(* IEC 61131-3 sources: ControlsBenchMUSE/codesys/library/source, 19 files *)

(* ---- ST_CB_Config.st ---- *)
TYPE ST_CB_Config :
STRUCT
    DomainId : UDINT; // nonzero; unique per authority domain in the application
    SchemaId : UDINT; // nonzero machine-map fingerprint of the raw channel layout
    TimeoutUs : ULINT := 500000; // heartbeat staleness as elapsed microseconds
    DigitalCount : UINT; // configured channels occupy indices 0..Count-1 of each bank
    SignedCount : UINT;
    UnsignedCount : UINT;
    RealCount : UINT;
    SignedBits : ARRAY[0..31] OF USINT; // native width of each configured channel: 8, 16 or 32
    UnsignedBits : ARRAY[0..31] OF USINT; // native width of each configured channel: 1 to 32
    RealNonFiniteAllowed : ARRAY[0..15] OF BOOL; // TRUE only where the device can report NaN or infinity
END_STRUCT
END_TYPE

(* ---- ST_CB_Image.st ---- *)
TYPE ST_CB_Image :
STRUCT
    Digital : ARRAY[0..63] OF BOOL;
    Numeric : ST_CB_Numeric;
END_STRUCT
END_TYPE

(* ---- ST_CB_ImageMask.st ---- *)
TYPE ST_CB_ImageMask :
STRUCT
    Digital : ARRAY[0..63] OF BOOL;
    Numeric : ST_CB_NumericMask;
END_STRUCT
END_TYPE

(* ---- ST_CB_Numeric.st ---- *)
TYPE ST_CB_Numeric :
STRUCT
    Signed : ARRAY[0..31] OF DINT;
    Unsigned : ARRAY[0..31] OF UDINT;
    RealValue : ARRAY[0..15] OF REAL;
END_STRUCT
END_TYPE

(* ---- ST_CB_NumericMask.st ---- *)
TYPE ST_CB_NumericMask :
STRUCT
    Signed : ARRAY[0..31] OF BOOL;
    Unsigned : ARRAY[0..31] OF BOOL;
    RealValue : ARRAY[0..15] OF BOOL;
END_STRUCT
END_TYPE

(* ---- ST_CB_ObservationFrame.st ---- *)
TYPE ST_CB_ObservationFrame :
STRUCT
    FrameFormat : UDINT := 1; // GVL_CB.FRAME_FORMAT_VERSION
    FrameSequence : ULINT; // frames published by this block since initialization
    BootIdentity : ULINT;
    DomainId : UDINT;
    SchemaId : UDINT;
    TapSchemaId : UDINT; // fingerprint of the configured tap list; 0 when none is configured
    SourceCycle : ULINT; // session cycle whose inputs and outputs this frame holds
    SourceTimeUs : ULINT; // platform monotonic time at capture, not wall-clock time
    CapturePhase : USINT; // GVL_CB.PHASE_POST_OUTPUT
    MissedCycles : ULINT; // cumulative session cycles that published no frame
    RepeatedCycles : ULINT; // cumulative calls without a new session cycle (integration error)
    SimApplied : BOOL; // SelectedInputs came from the workstation, not hardware
    ConnectorStale : BOOL;
    ConfigValid : BOOL;
    ClockValid : BOOL;
    ReconfigureRequired : BOOL;
    AnySuppressed : BOOL;
    AppliedEpoch : ULINT;
    AppliedSequence : ULINT;
    RawInputs : ST_CB_Image; // hardware values presented to the session, in either mode
    SelectedInputs : ST_CB_Image; // image the application consumed
    Commands : ST_CB_Image; // authentic application commands before suppression
    Physical : ST_CB_Image; // physical sink values after suppression
    Suppressed : ST_CB_ImageMask; // channels whose physical sink was suppressed
    Taps : ST_CB_Image; // explicitly configured observation taps; never writable through this library
END_STRUCT
END_TYPE

(* ---- ST_CB_Request.st ---- *)
TYPE ST_CB_Request :
STRUCT
    SimRequest : BOOL;
    SimulationResetRequest : BOOL; // rising edge: zero image, remain simulated
    SessionResetRequest : BOOL;
    Heartbeat : ULINT;
    RequestedSlot : USINT := 255;
    RequestedEpoch : ULINT;
    RequestedSequence : ULINT; // write LAST after validity/payload/metadata
    Slots : ARRAY[0..1] OF ST_CB_Slot;
END_STRUCT
END_TYPE

(* ---- ST_CB_Slot.st ---- *)
TYPE ST_CB_Slot :
STRUCT
    Valid : BOOL;
    DomainId : UDINT;
    SchemaId : UDINT;
    Epoch : ULINT;
    Sequence : ULINT;
    Data : ST_CB_Image;
END_STRUCT
END_TYPE

(* ---- ST_CB_Status.st ---- *)
TYPE ST_CB_Status :
STRUCT
    ProtocolVersion : UDINT := 2; // GVL_CB.PROTOCOL_VERSION
    DomainId : UDINT; // pinned at initialization
    SchemaId : UDINT; // pinned at initialization
    ConfigValid : BOOL;
    ClockValid : BOOL; // this cycle's time was not earlier than the previous cycle's
    ReconfigureRequired : BOOL; // latched by config, boot or clock change; cleared only by Reinitialize
    SimApplied : BOOL; // TRUE: the application consumes the workstation image
    ConnectorStale : BOOL := TRUE;
    BootIdentity : ULINT;
    Cycle : ULINT; // calls of this domain session, not universal PLC scans
    TimeUs : ULINT;
    LastHeartbeat : ULINT;
    LastHeartbeatTimeUs : ULINT;
    ActiveSlot : USINT := 255;
    AppliedEpoch : ULINT;
    AppliedSequence : ULINT;
    AppliedCycle : ULINT;
    AppliedTimeUs : ULINT;
    // Acknowledgement of the last consumed request event, accepted or not.
    ConsumedEpoch : ULINT;
    ConsumedSequence : ULINT;
    ConsumedSlot : USINT := 255;
    ConsumedResult : UINT; // GVL_CB.RESULT_*
    ConsumedCycle : ULINT;
    ConsumedTimeUs : ULINT;
    RejectBank : USINT; // GVL_CB.BANK_* of the first channel failing representation checks
    RejectIndex : UINT;
    CommitCount : ULINT;
    DuplicateCount : ULINT;
    StaleCount : ULINT;
    SkippedCount : ULINT;
    InvalidSlotCount : ULINT;
    IncompleteSlotCount : ULINT;
    MetadataMismatchCount : ULINT;
    RepresentationRejectedCount : ULINT;
    EpochRejectedCount : ULINT;
    NotSimulatedCount : ULINT;
    BlockedRequestCount : ULINT;
    IdleClearCount : ULINT;
    SessionResetCount : ULINT;
    SimulationResetCount : ULINT;
    SimulationEntryCount : ULINT;
    ReinitializeCount : ULINT;
END_STRUCT
END_TYPE

(* ---- U_CB_Real32.st ---- *)
TYPE U_CB_Real32 :
UNION
    AsReal : REAL; // IEEE 754 binary32 value
    AsBits : DWORD; // the same 32 bits, for encoding checks without numeric conversion
END_UNION
END_TYPE

(* ---- GVL_CB.st ---- *)
{attribute 'qualified_only'}
VAR_GLOBAL CONSTANT
    // Interface versions. The package version is the library project version (VERSIONING.md).
    API_VERSION_MAJOR : UINT := 0;
    API_VERSION_MINOR : UINT := 2;
    PROTOCOL_VERSION : UDINT := 2; // request, slot and status semantics of this raw-bank profile
    FRAME_FORMAT_VERSION : UDINT := 1; // ST_CB_ObservationFrame layout and meaning
    // Fixed capacities of ST_CB_Image. Configured channels occupy indices 0..Count-1.
    DIGITAL_CAPACITY : UINT := 64;
    SIGNED_CAPACITY : UINT := 32;
    UNSIGNED_CAPACITY : UINT := 32;
    REAL_CAPACITY : UINT := 16;
    NO_SLOT : USINT := 255;
    // Status.ConsumedResult: outcome of the last request event the session consumed.
    RESULT_NONE : UINT := 0;
    RESULT_ACCEPTED : UINT := 1;
    RESULT_IDLE_CLEARED : UINT := 2;
    RESULT_INVALID_SLOT : UINT := 3;
    RESULT_INCOMPLETE_SLOT : UINT := 4;
    RESULT_METADATA_MISMATCH : UINT := 5;
    RESULT_DUPLICATE : UINT := 6;
    RESULT_STALE : UINT := 7;
    RESULT_EPOCH_REJECTED : UINT := 8;
    RESULT_REPRESENTATION : UINT := 9;
    RESULT_NOT_SIMULATED : UINT := 10;
    RESULT_CONFIG_INVALID : UINT := 11;
    RESULT_RECONFIGURE_REQUIRED : UINT := 12;
    RESULT_SESSION_RESET : UINT := 13;
    RESULT_SIMULATION_RESET : UINT := 14;
    RESULT_SIMULATION_ENTRY : UINT := 15;
    RESULT_REINITIALIZED : UINT := 16;
    // Status.RejectBank: bank of the first channel that failed representation checks.
    BANK_NONE : USINT := 0;
    BANK_DIGITAL : USINT := 1;
    BANK_SIGNED : USINT := 2;
    BANK_UNSIGNED : USINT := 3;
    BANK_REAL : USINT := 4;
    // ST_CB_ObservationFrame.CapturePhase.
    PHASE_POST_OUTPUT : USINT := 2;
END_VAR

(* ---- F_CB_CheckImage.st ---- *)
FUNCTION F_CB_CheckImage : UINT
VAR_INPUT
    Image : ST_CB_Image; // candidate image from a workstation slot
    Config : ST_CB_Config; // pinned domain configuration
END_VAR
VAR_OUTPUT
    Bank : USINT; // GVL_CB.BANK_* of the first failing channel
    Index : UINT;
END_VAR
VAR
    i : UINT;
    bits : USINT;
    maxValue : UDINT;
    raw : U_CB_Real32;
END_VAR
// Rejects values a configured native type cannot represent, non-finite REAL on
// finite-only channels, and nonzero data in unconfigured channels. It never
// clamps, rounds or substitutes a value; the caller keeps the prior image.
F_CB_CheckImage := GVL_CB.RESULT_NONE;
Bank := GVL_CB.BANK_NONE;
Index := 0;
FOR i := 0 TO 63 DO
    IF (i >= Config.DigitalCount) AND Image.Digital[i] THEN
        F_CB_CheckImage := GVL_CB.RESULT_REPRESENTATION;
        Bank := GVL_CB.BANK_DIGITAL;
        Index := i;
        RETURN;
    END_IF;
END_FOR;
FOR i := 0 TO 31 DO
    IF i < Config.SignedCount THEN
        bits := Config.SignedBits[i];
        IF ((bits = 8) AND ((Image.Numeric.Signed[i] < -128) OR (Image.Numeric.Signed[i] > 127)))
            OR ((bits = 16) AND ((Image.Numeric.Signed[i] < -32768) OR (Image.Numeric.Signed[i] > 32767))) THEN
            F_CB_CheckImage := GVL_CB.RESULT_REPRESENTATION;
            Bank := GVL_CB.BANK_SIGNED;
            Index := i;
            RETURN;
        END_IF;
    ELSIF Image.Numeric.Signed[i] <> 0 THEN
        F_CB_CheckImage := GVL_CB.RESULT_REPRESENTATION;
        Bank := GVL_CB.BANK_SIGNED;
        Index := i;
        RETURN;
    END_IF;
END_FOR;
FOR i := 0 TO 31 DO
    IF i < Config.UnsignedCount THEN
        bits := Config.UnsignedBits[i];
        IF bits >= 32 THEN
            maxValue := 16#FFFFFFFF;
        ELSE
            maxValue := SHL(UDINT#1, bits) - 1;
        END_IF;
        IF Image.Numeric.Unsigned[i] > maxValue THEN
            F_CB_CheckImage := GVL_CB.RESULT_REPRESENTATION;
            Bank := GVL_CB.BANK_UNSIGNED;
            Index := i;
            RETURN;
        END_IF;
    ELSIF Image.Numeric.Unsigned[i] <> 0 THEN
        F_CB_CheckImage := GVL_CB.RESULT_REPRESENTATION;
        Bank := GVL_CB.BANK_UNSIGNED;
        Index := i;
        RETURN;
    END_IF;
END_FOR;
FOR i := 0 TO 15 DO
    raw.AsReal := Image.Numeric.RealValue[i];
    IF i < Config.RealCount THEN
        IF ((raw.AsBits AND 16#7F800000) = 16#7F800000) AND NOT Config.RealNonFiniteAllowed[i] THEN
            F_CB_CheckImage := GVL_CB.RESULT_REPRESENTATION;
            Bank := GVL_CB.BANK_REAL;
            Index := i;
            RETURN;
        END_IF;
    ELSIF raw.AsBits <> 0 THEN
        F_CB_CheckImage := GVL_CB.RESULT_REPRESENTATION;
        Bank := GVL_CB.BANK_REAL;
        Index := i;
        RETURN;
    END_IF;
END_FOR;
END_FUNCTION

(* ---- FB_CB_AI.st ---- *)
FUNCTION_BLOCK FB_CB_AI
VAR_INPUT
    Hardware : ST_CB_Numeric;
    Simulated : ST_CB_Numeric;
    SimApplied : BOOL;
END_VAR
VAR_OUTPUT
    Selected : ST_CB_Numeric;
END_VAR
IF SimApplied THEN Selected := Simulated; ELSE Selected := Hardware; END_IF;
END_FUNCTION_BLOCK

(* ---- FB_CB_AO.st ---- *)
FUNCTION_BLOCK FB_CB_AO
VAR_INPUT
    Commands : ST_CB_Numeric; // authentic application commands
    Suppress : ST_CB_NumericMask; // explicit physical-sink configuration
    SuppressedValues : ST_CB_Numeric; // physical value while suppressed; default raw zero
END_VAR
VAR_OUTPUT
    Observed : ST_CB_Numeric; // always the authentic commands
    Physical : ST_CB_Numeric; // value for the physical sink
    Applied : ST_CB_NumericMask; // suppression mask applied by this call
    SuppressedCount : UINT;
END_VAR
VAR
    i : UINT;
END_VAR
Observed := Commands;
Physical := Commands;
Applied := Suppress;
SuppressedCount := 0;
FOR i := 0 TO 31 DO
    IF Suppress.Signed[i] THEN
        Physical.Signed[i] := SuppressedValues.Signed[i];
        SuppressedCount := SuppressedCount + 1;
    END_IF;
    IF Suppress.Unsigned[i] THEN
        Physical.Unsigned[i] := SuppressedValues.Unsigned[i];
        SuppressedCount := SuppressedCount + 1;
    END_IF;
END_FOR;
FOR i := 0 TO 15 DO
    IF Suppress.RealValue[i] THEN
        Physical.RealValue[i] := SuppressedValues.RealValue[i];
        SuppressedCount := SuppressedCount + 1;
    END_IF;
END_FOR;
END_FUNCTION_BLOCK

(* ---- FB_CB_DI.st ---- *)
FUNCTION_BLOCK FB_CB_DI
VAR_INPUT
    Hardware : ARRAY[0..63] OF BOOL;
    Simulated : ARRAY[0..63] OF BOOL;
    SimApplied : BOOL;
END_VAR
VAR_OUTPUT
    Selected : ARRAY[0..63] OF BOOL;
END_VAR
IF SimApplied THEN Selected := Simulated; ELSE Selected := Hardware; END_IF;
END_FUNCTION_BLOCK

(* ---- FB_CB_DO.st ---- *)
FUNCTION_BLOCK FB_CB_DO
VAR_INPUT
    Commands : ARRAY[0..63] OF BOOL; // authentic application commands
    Suppress : ARRAY[0..63] OF BOOL; // explicit physical-sink configuration
    SuppressedValues : ARRAY[0..63] OF BOOL; // physical value while suppressed; default FALSE
END_VAR
VAR_OUTPUT
    Observed : ARRAY[0..63] OF BOOL; // always the authentic commands
    Physical : ARRAY[0..63] OF BOOL; // value for the physical sink
    Applied : ARRAY[0..63] OF BOOL; // suppression mask applied by this call
    SuppressedCount : UINT;
END_VAR
VAR
    i : UINT;
END_VAR
Observed := Commands;
Applied := Suppress;
SuppressedCount := 0;
FOR i := 0 TO 63 DO
    IF Suppress[i] THEN
        Physical[i] := SuppressedValues[i];
        SuppressedCount := SuppressedCount + 1;
    ELSE
        Physical[i] := Commands[i];
    END_IF;
END_FOR;
END_FUNCTION_BLOCK

(* ---- FB_CB_Observation.st ---- *)
FUNCTION_BLOCK FB_CB_Observation
VAR_INPUT
    Enable : BOOL := TRUE; // FALSE keeps the last frame; the gap is counted when re-enabled
    InputStatus : ST_CB_Status; // Status of the same domain session, this cycle
    RawInputs : ST_CB_Image; // the Hardware image given to the session this cycle
    SelectedInputs : ST_CB_Image; // the session Image the application consumed
    Commands : ST_CB_Image; // authentic commands, before suppression
    Physical : ST_CB_Image; // physical sink values, after suppression
    Suppressed : ST_CB_ImageMask; // applied suppression masks from the DO/AO taps
    Taps : ST_CB_Image; // explicitly configured observation taps packed by the machine map
    TapSchemaId : UDINT; // tap-list fingerprint from the machine map; 0 when none is configured
    NowUs : ULINT;
END_VAR
VAR_OUTPUT
    PublicationRevision : ULINT; // odd while updating; even after publication
    Frame : ST_CB_ObservationFrame;
END_VAR
VAR
    haveCycle : BOOL;
    lastCycle : ULINT;
    anySuppressed : BOOL;
    i : UINT;
END_VAR
// Passive observation: needs no simulation authority or suppression and writes
// nothing back. Call once per cycle after the output taps, in the session's task.
// Fixed-size copy, no allocation, no waiting on any transport.
IF NOT Enable THEN
    RETURN;
END_IF;
anySuppressed := FALSE;
FOR i := 0 TO 63 DO
    anySuppressed := anySuppressed OR Suppressed.Digital[i];
END_FOR;
FOR i := 0 TO 31 DO
    anySuppressed := anySuppressed OR Suppressed.Numeric.Signed[i] OR Suppressed.Numeric.Unsigned[i];
END_FOR;
FOR i := 0 TO 15 DO
    anySuppressed := anySuppressed OR Suppressed.Numeric.RealValue[i];
END_FOR;
PublicationRevision := PublicationRevision + 1;
IF haveCycle THEN
    IF InputStatus.Cycle = lastCycle THEN
        Frame.RepeatedCycles := Frame.RepeatedCycles + 1;
    ELSIF InputStatus.Cycle > lastCycle + 1 THEN
        Frame.MissedCycles := Frame.MissedCycles + (InputStatus.Cycle - lastCycle - 1);
    END_IF;
END_IF;
haveCycle := TRUE;
lastCycle := InputStatus.Cycle;
Frame.FrameFormat := GVL_CB.FRAME_FORMAT_VERSION;
Frame.FrameSequence := Frame.FrameSequence + 1;
Frame.BootIdentity := InputStatus.BootIdentity;
Frame.DomainId := InputStatus.DomainId;
Frame.SchemaId := InputStatus.SchemaId;
Frame.TapSchemaId := TapSchemaId;
Frame.SourceCycle := InputStatus.Cycle;
Frame.SourceTimeUs := NowUs;
Frame.CapturePhase := GVL_CB.PHASE_POST_OUTPUT;
Frame.SimApplied := InputStatus.SimApplied;
Frame.ConnectorStale := InputStatus.ConnectorStale;
Frame.ConfigValid := InputStatus.ConfigValid;
Frame.ClockValid := InputStatus.ClockValid;
Frame.ReconfigureRequired := InputStatus.ReconfigureRequired;
Frame.AnySuppressed := anySuppressed;
Frame.AppliedEpoch := InputStatus.AppliedEpoch;
Frame.AppliedSequence := InputStatus.AppliedSequence;
Frame.RawInputs := RawInputs;
Frame.SelectedInputs := SelectedInputs;
Frame.Commands := Commands;
Frame.Physical := Physical;
Frame.Suppressed := Suppressed;
Frame.Taps := Taps;
PublicationRevision := PublicationRevision + 1;
END_FUNCTION_BLOCK

(* ---- FB_CB_OutputCapture.st ---- *)
FUNCTION_BLOCK FB_CB_OutputCapture
VAR_INPUT
    InputStatus : ST_CB_Status;
    Commands : ST_CB_Image;
    NowUs : ULINT;
END_VAR
VAR_OUTPUT
    PublicationRevision : ULINT; // odd while updating; even after publication
    Observed : ST_CB_Image;
    BootIdentity : ULINT;
    DomainId : UDINT;
    SchemaId : UDINT;
    SourceSimulated : BOOL;
    SourceEpoch : ULINT;
    SourceSequence : ULINT;
    InputAppliedCycle : ULINT;
    CaptureCycle : ULINT;
    CaptureTimeUs : ULINT;
END_VAR
// Call after application/output computation, within the same task as Session.
PublicationRevision := PublicationRevision + 1;
Observed := Commands;
BootIdentity := InputStatus.BootIdentity;
DomainId := InputStatus.DomainId;
SchemaId := InputStatus.SchemaId;
SourceSimulated := InputStatus.SimApplied;
SourceEpoch := InputStatus.AppliedEpoch;
SourceSequence := InputStatus.AppliedSequence;
InputAppliedCycle := InputStatus.AppliedCycle;
CaptureCycle := InputStatus.Cycle;
CaptureTimeUs := NowUs;
PublicationRevision := PublicationRevision + 1;
END_FUNCTION_BLOCK

(* ---- FB_CB_Session.st ---- *)
FUNCTION_BLOCK FB_CB_Session
VAR_INPUT
    Hardware : ST_CB_Image; // raw values packed by the machine mapping, unchanged
    Config : ST_CB_Config; // pinned at initialization; any later change latches ReconfigureRequired
    NowUs : ULINT; // monotonic microseconds from a platform service
    BootId : ULINT; // nonzero platform identity that changes on every application or runtime restart
    Reinitialize : BOOL; // rising edge from local application authority, never from the workstation
END_VAR
VAR_IN_OUT
    Request : ST_CB_Request; // storage owned by this domain; exactly one workstation writer
END_VAR
VAR_OUTPUT
    Image : ST_CB_Image; // complete image the application consumes this cycle
    Status : ST_CB_Status;
END_VAR
VAR
    initialized : BOOL;
    previousSim : BOOL;
    previousSessionReset : BOOL;
    previousSimulationReset : BOOL;
    previousReinitialize : BOOL;
    haveHeartbeat : BOOL;
    previousHeartbeat : ULINT;
    lastHeartbeatUs : ULINT;
    lastTimeUs : ULINT;
    lastRequestSequence : ULINT;
    active : ST_CB_Image;
    zero : ST_CB_Image;
    pinned : ST_CB_Config;
    slot : ST_CB_Slot;
    reqSim : BOOL;
    reqSessionReset : BOOL;
    reqSimulationReset : BOOL;
    reqHeartbeat : ULINT;
    reqSlot : USINT;
    reqEpoch : ULINT;
    reqSequence : ULINT;
    reinitializeEdge : BOOL;
    entryEdge : BOOL;
    sessionResetEdge : BOOL;
    simulationResetEdge : BOOL;
    commitEdge : BOOL;
    configChanged : BOOL;
    blocked : BOOL;
    blockedResult : UINT;
    staleAtEntry : BOOL;
    accept : BOOL;
    consumed : BOOL;
    result : UINT;
    rejectBank : USINT;
    rejectIndex : UINT;
    i : UINT;
    di : FB_CB_DI;
    ai : FB_CB_AI;
END_VAR
// Read each request word once so every decision in this cycle uses the same values.
reqSim := Request.SimRequest;
reqSessionReset := Request.SessionResetRequest;
reqSimulationReset := Request.SimulationResetRequest;
reqHeartbeat := Request.Heartbeat;
reqSlot := Request.RequestedSlot;
reqEpoch := Request.RequestedEpoch;
reqSequence := Request.RequestedSequence;
consumed := FALSE;
result := GVL_CB.RESULT_NONE;
reinitializeEdge := Reinitialize AND NOT previousReinitialize;
previousReinitialize := Reinitialize;
Status.Cycle := Status.Cycle + 1;
Status.TimeUs := NowUs;

IF NOT initialized OR reinitializeEdge THEN
    // A fresh domain pins configuration and boot identity, holds raw zero and
    // consumes whatever is staged; a heartbeat must change before the link is fresh.
    pinned := Config;
    Status.BootIdentity := BootId;
    Status.ReconfigureRequired := FALSE;
    active := zero;
    Status.ActiveSlot := GVL_CB.NO_SLOT;
    Status.AppliedEpoch := 0;
    Status.AppliedSequence := 0;
    Status.AppliedCycle := Status.Cycle;
    Status.AppliedTimeUs := NowUs;
    lastTimeUs := NowUs;
    lastRequestSequence := reqSequence;
    previousHeartbeat := reqHeartbeat;
    haveHeartbeat := FALSE;
    IF initialized THEN
        previousSim := reqSim; // a simulated domain stays simulated, now at raw zero
        Status.ReinitializeCount := Status.ReinitializeCount + 1;
        consumed := TRUE;
        result := GVL_CB.RESULT_REINITIALIZED;
    END_IF;
    initialized := TRUE;
END_IF;
Status.DomainId := pinned.DomainId;
Status.SchemaId := pinned.SchemaId;

// Configuration validity: identities, capacities and declared native widths.
Status.ConfigValid := (Config.DomainId <> 0) AND (Config.SchemaId <> 0) AND (Config.TimeoutUs > 0)
    AND (Config.DigitalCount <= GVL_CB.DIGITAL_CAPACITY) AND (Config.SignedCount <= GVL_CB.SIGNED_CAPACITY)
    AND (Config.UnsignedCount <= GVL_CB.UNSIGNED_CAPACITY) AND (Config.RealCount <= GVL_CB.REAL_CAPACITY)
    AND (BootId <> 0);
configChanged := (Config.DomainId <> pinned.DomainId) OR (Config.SchemaId <> pinned.SchemaId)
    OR (Config.TimeoutUs <> pinned.TimeoutUs) OR (Config.DigitalCount <> pinned.DigitalCount)
    OR (Config.SignedCount <> pinned.SignedCount) OR (Config.UnsignedCount <> pinned.UnsignedCount)
    OR (Config.RealCount <> pinned.RealCount);
FOR i := 0 TO 31 DO
    IF (i < Config.SignedCount) AND NOT ((Config.SignedBits[i] = 8) OR (Config.SignedBits[i] = 16)
        OR (Config.SignedBits[i] = 32)) THEN
        Status.ConfigValid := FALSE;
    END_IF;
    IF (i < Config.UnsignedCount) AND ((Config.UnsignedBits[i] = 0) OR (Config.UnsignedBits[i] > 32)) THEN
        Status.ConfigValid := FALSE;
    END_IF;
    IF (Config.SignedBits[i] <> pinned.SignedBits[i]) OR (Config.UnsignedBits[i] <> pinned.UnsignedBits[i]) THEN
        configChanged := TRUE;
    END_IF;
END_FOR;
FOR i := 0 TO 15 DO
    IF Config.RealNonFiniteAllowed[i] <> pinned.RealNonFiniteAllowed[i] THEN
        configChanged := TRUE;
    END_IF;
END_FOR;
Status.ClockValid := NowUs >= lastTimeUs;
IF configChanged OR (BootId <> Status.BootIdentity) OR NOT Status.ClockValid THEN
    Status.ReconfigureRequired := TRUE; // no hidden remapping; Reinitialize explicitly
END_IF;
blocked := NOT Status.ConfigValid OR Status.ReconfigureRequired;
IF Status.ReconfigureRequired THEN
    blockedResult := GVL_CB.RESULT_RECONFIGURE_REQUIRED;
ELSE
    blockedResult := GVL_CB.RESULT_CONFIG_INVALID;
END_IF;

// Link freshness uses elapsed microseconds, independent of the task period.
// Staleness at cycle entry is evaluated before this cycle's heartbeat is applied.
staleAtEntry := NOT haveHeartbeat OR (NowUs < lastHeartbeatUs)
    OR ((NowUs - lastHeartbeatUs) > pinned.TimeoutUs);
IF reqHeartbeat <> previousHeartbeat THEN
    previousHeartbeat := reqHeartbeat;
    lastHeartbeatUs := NowUs;
    haveHeartbeat := TRUE;
    Status.LastHeartbeat := reqHeartbeat;
    Status.LastHeartbeatTimeUs := NowUs;
END_IF;
Status.ConnectorStale := NOT haveHeartbeat OR (NowUs < lastHeartbeatUs)
    OR ((NowUs - lastHeartbeatUs) > pinned.TimeoutUs);

entryEdge := reqSim AND NOT previousSim;
previousSim := reqSim;
sessionResetEdge := reqSessionReset AND NOT previousSessionReset;
previousSessionReset := reqSessionReset;
simulationResetEdge := reqSimulationReset AND NOT previousSimulationReset;
previousSimulationReset := reqSimulationReset;
commitEdge := reqSequence <> lastRequestSequence;

IF entryEdge THEN
    // Entry gives the workstation complete input authority at raw zero.
    // Staged data never applies on entry; complete commits establish normal conditions.
    active := zero;
    Status.ActiveSlot := GVL_CB.NO_SLOT;
    Status.AppliedEpoch := 0;
    Status.AppliedSequence := 0;
    Status.AppliedCycle := Status.Cycle;
    Status.AppliedTimeUs := NowUs;
    Status.SimulationEntryCount := Status.SimulationEntryCount + 1;
    consumed := TRUE;
    result := GVL_CB.RESULT_SIMULATION_ENTRY;
    lastRequestSequence := reqSequence;
    commitEdge := FALSE;
END_IF;

IF simulationResetEdge OR sessionResetEdge THEN
    // Neither reset requests a machine Reset or leaves simulation.
    IF blocked THEN
        Status.BlockedRequestCount := Status.BlockedRequestCount + 1;
        result := blockedResult;
    ELSE
        IF simulationResetEdge THEN
            active := zero; // explicit simulation reset: raw zero, still simulated
            Status.SimulationResetCount := Status.SimulationResetCount + 1;
            result := GVL_CB.RESULT_SIMULATION_RESET;
        END_IF;
        IF sessionResetEdge THEN
            Status.SessionResetCount := Status.SessionResetCount + 1; // image retained
            IF NOT simulationResetEdge THEN
                result := GVL_CB.RESULT_SESSION_RESET;
            END_IF;
        END_IF;
        Status.ActiveSlot := GVL_CB.NO_SLOT;
        Status.AppliedEpoch := 0;
        Status.AppliedSequence := 0;
        Status.AppliedCycle := Status.Cycle;
        Status.AppliedTimeUs := NowUs;
    END_IF;
    consumed := TRUE;
    lastRequestSequence := reqSequence; // the staged request is consumed without applying
    commitEdge := FALSE;
END_IF;

IF commitEdge THEN
    // RequestedSequence, written last, is the single commit edge. Each edge is consumed once.
    consumed := TRUE;
    accept := FALSE;
    rejectBank := GVL_CB.BANK_NONE;
    rejectIndex := 0;
    IF blocked THEN
        Status.BlockedRequestCount := Status.BlockedRequestCount + 1;
        result := blockedResult;
    ELSIF NOT reqSim THEN
        Status.NotSimulatedCount := Status.NotSimulatedCount + 1;
        result := GVL_CB.RESULT_NOT_SIMULATED;
    ELSIF (reqEpoch = 0) AND (reqSequence = 0) THEN
        Status.IdleClearCount := Status.IdleClearCount + 1;
        result := GVL_CB.RESULT_IDLE_CLEARED;
    ELSIF (reqSlot > 1) OR (reqSlot = Status.ActiveSlot) THEN
        Status.InvalidSlotCount := Status.InvalidSlotCount + 1;
        result := GVL_CB.RESULT_INVALID_SLOT;
    ELSE
        slot := Request.Slots[reqSlot];
        IF NOT slot.Valid OR (slot.Epoch = 0) OR (slot.Sequence = 0) THEN
            Status.IncompleteSlotCount := Status.IncompleteSlotCount + 1;
            result := GVL_CB.RESULT_INCOMPLETE_SLOT;
        ELSIF (slot.DomainId <> pinned.DomainId) OR (slot.SchemaId <> pinned.SchemaId)
            OR (slot.Epoch <> reqEpoch) OR (slot.Sequence <> reqSequence) THEN
            Status.MetadataMismatchCount := Status.MetadataMismatchCount + 1;
            result := GVL_CB.RESULT_METADATA_MISMATCH;
        ELSE
            result := F_CB_CheckImage(Image := slot.Data, Config := pinned, Bank => rejectBank, Index => rejectIndex);
            IF result <> GVL_CB.RESULT_NONE THEN
                Status.RepresentationRejectedCount := Status.RepresentationRejectedCount + 1;
            ELSIF Status.AppliedEpoch = 0 THEN
                accept := TRUE;
            ELSIF slot.Epoch = Status.AppliedEpoch THEN
                IF slot.Sequence = Status.AppliedSequence THEN
                    Status.DuplicateCount := Status.DuplicateCount + 1;
                    result := GVL_CB.RESULT_DUPLICATE;
                ELSIF slot.Sequence < Status.AppliedSequence THEN
                    Status.StaleCount := Status.StaleCount + 1;
                    result := GVL_CB.RESULT_STALE;
                ELSE
                    IF slot.Sequence - Status.AppliedSequence > 1 THEN
                        Status.SkippedCount := Status.SkippedCount + 1;
                    END_IF;
                    accept := TRUE;
                END_IF;
            ELSIF staleAtEntry THEN
                accept := TRUE; // a new epoch only after elapsed staleness or an explicit reset
            ELSE
                Status.EpochRejectedCount := Status.EpochRejectedCount + 1;
                result := GVL_CB.RESULT_EPOCH_REJECTED;
            END_IF;
        END_IF;
    END_IF;
    IF accept THEN
        active := slot.Data; // every bank changes together; no torn image
        Status.ActiveSlot := reqSlot;
        Status.AppliedEpoch := slot.Epoch;
        Status.AppliedSequence := slot.Sequence;
        Status.AppliedCycle := Status.Cycle;
        Status.AppliedTimeUs := NowUs;
        Status.CommitCount := Status.CommitCount + 1;
        result := GVL_CB.RESULT_ACCEPTED;
    END_IF;
    Status.RejectBank := rejectBank;
    Status.RejectIndex := rejectIndex;
    lastRequestSequence := reqSequence;
END_IF;

IF consumed THEN
    Status.ConsumedEpoch := reqEpoch;
    Status.ConsumedSequence := reqSequence;
    Status.ConsumedSlot := reqSlot;
    Status.ConsumedResult := result;
    Status.ConsumedCycle := Status.Cycle;
    Status.ConsumedTimeUs := NowUs;
END_IF;

// Exit Simulation (SimRequest FALSE) is always honoured. Bad configuration while
// simulated holds the image; it never silently selects hardware.
Status.SimApplied := reqSim;
di(Hardware := Hardware.Digital, Simulated := active.Digital, SimApplied := reqSim);
ai(Hardware := Hardware.Numeric, Simulated := active.Numeric, SimApplied := reqSim);
Image.Digital := di.Selected;
Image.Numeric := ai.Selected;
lastTimeUs := NowUs;
END_FUNCTION_BLOCK
